TYPE ST_AlarmRef :
STRUCT
	stControl					:ST_AlarmOut;
	stManual					:ST_AlarmOut;
	stMaintenance			:ST_AlarmOut;
	stHome					:ST_AlarmOut;
	stAuto					:ST_AlarmOut;
END_STRUCT
END_TYPE

(* stored: Version 1.1.0.1, ProductVersion 3.1.4024.15
   DUT ST_AlarmRef: Id {99efbea5-b2bb-4a78-9560-ebb4fad806f9} *)
